// SIMATIC S7-200 project (STEP 7-Micro/WIN), CPU 224XP CN REL 02.01

SYMBOL_TABLE USUARIO1
SO               I0.3     // Sensor de Objetos (Detecta la pieza para iniciar la seleccion)
S_I              I0.4     // Sensor de fibra Optica (clasificacion de materiales)
SM               I0.5     // Sensor magnetico (clasificacion de materiales)
S1               I0.7     // Sensor de retorno del cilindro 1
S2               I1.0     // Sensor de retorno del cilindro 2
S3               I1.1     // Sensor de retorno del cilindro 3
SBB1             I1.3     // Pulsador de Marcha
SBB2             I1.2     // Pulsador de Paro
QS               I1.4     // Zeta de emergencia
SA               I1.5     // Selector rotatorio
am               Q0.0     // Motor
C_1              Q0.4     // cilindro neumatico 1
C_2              Q0.5     // cilindro neumatico 2
C_3              Q0.6     // cilindro neumatico 3
HL1              Q0.7     // Lampara de señalizacion amarilla
HL2              Q1.0     // Lampara de señalizacion verde
HL3              Q1.1     // Lampara de señalizacion roja
E0               M0.0     // Estado 0
E1               M0.1     // Estado 1
E2               M0.2     // Estado 2
E3               M0.3     // Estado 3
E4               M0.4     // Estado 4
E5               M0.5     // Estado 5
E6               M0.6     // Estado 6
E7               M0.7     // Estado 7
E8               M1.0     // Estado 8
E9               M1.1     // Estado 9
E10              M1.2     // Estado 10
E11              M1.3     // Estado 11
E12              M1.4     // Estado 12
E13              M1.5     // Estado 13
E14              M1.6     // Estado 14
EM               M1.7     // Variable para paro momentaneo
MOTOR            M2.0     // Variable para activacion o desactivacion del motor
E15              M2.1     // Estado 15
E16              M2.2     // Estado 16
C_c1             VD100
C_0              VD110
y_k              VD180
r_k              VD190
u_k              VD120
xh1_k_1          VD130
xh1_k            VD140
xh2_k_1          VD300
xh2_k            VD160
xh3_k_1          VD170
xh3_k            VD200
xp1_k            VD210
xp2_k            VD220
xp3_k            VD230
Ao               VD310
Bo               VD320
Co               VD330
Do               VD340
Eo               VD350
Fo               VD360
Go               VD370
Ho               VD380
Io               VD390
Jo               VD400
L1o              VD410
L2o              VD420
L3o              VD430
e_k              VD270
Ee               VD240
r_k_1            VD250
u_k_1            VD150
k1o              VD440
k2o              VD450
k3o              VD460
END_SYMBOL_TABLE

ORGANIZATION_BLOCK PRINCIPAL:OB1
TITLE=UNIDAD DE SELECCION
BEGIN
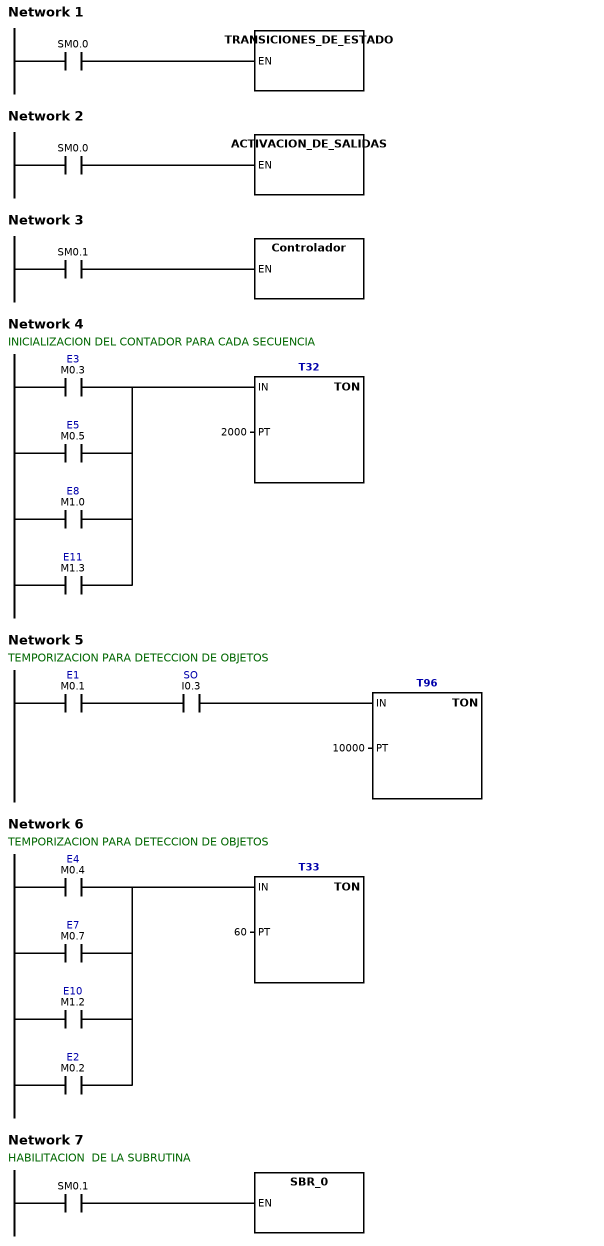
Network 1
LD     SM0.0
CALL   TRANSICIONES_DE_ESTADO:SBR1
Network 2
LD     SM0.0
CALL   ACTIVACION_DE_SALIDAS:SBR2
Network 3
LD     SM0.1
CALL   Controlador:SBR3
Network 4
// INICIALIZACION DEL CONTADOR PARA CADA SECUENCIA 
LD     E3:M0.3
O      E5:M0.5
O      E8:M1.0
O      E11:M1.3
TON    T32, 2000
Network 5
// TEMPORIZACION PARA DETECCION DE OBJETOS
LD     E1:M0.1
A      SO:I0.3
TON    T96, 10000
Network 6
// TEMPORIZACION PARA DETECCION DE OBJETOS
LD     E4:M0.4
O      E7:M0.7
O      E10:M1.2
O      E2:M0.2
TON    T33, 60
Network 7
// HABILITACION  DE LA SUBRUTINA
LD     SM0.1
CALL   SBR_0:SBR0
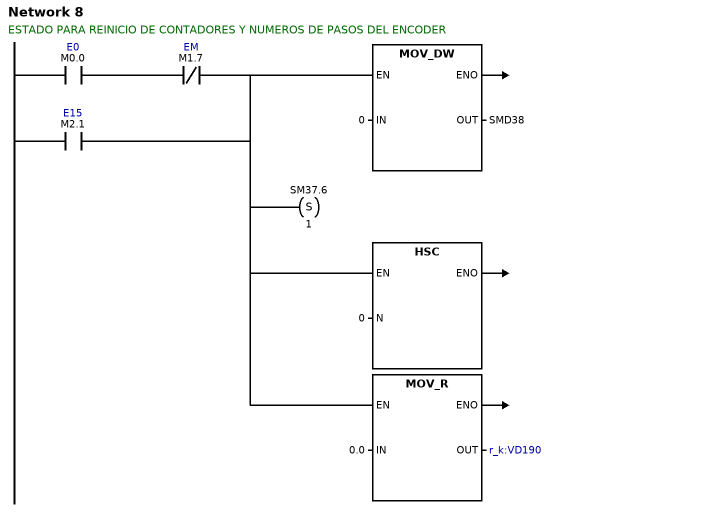
Network 8
// ESTADO PARA REINICIO DE CONTADORES Y NUMEROS DE PASOS DEL ENCODER
LD     E0:M0.0
AN     EM:M1.7
O      E15:M2.1
MOVD   0, SMD38
S      SM37.6, 1
HSC    0
MOVR   0.0, r_k:VD190
END_ORGANIZATION_BLOCK

SUBROUTINE_BLOCK SBR_0:SBR0
TITLE=COMENTARIOS DE LA SUBRUTINA
BEGIN
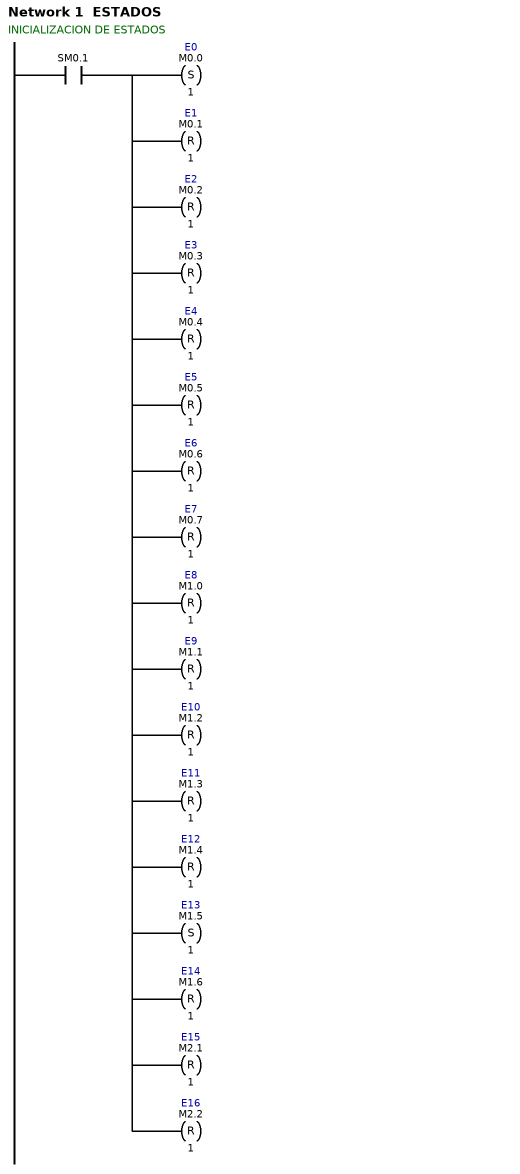
Network 1 // ESTADOS
// INICIALIZACION DE ESTADOS
LD     SM0.1
S      E0:M0.0, 1
R      E1:M0.1, 1
R      E2:M0.2, 1
R      E3:M0.3, 1
R      E4:M0.4, 1
R      E5:M0.5, 1
R      E6:M0.6, 1
R      E7:M0.7, 1
R      E8:M1.0, 1
R      E9:M1.1, 1
R      E10:M1.2, 1
R      E11:M1.3, 1
R      E12:M1.4, 1
S      E13:M1.5, 1
R      E14:M1.6, 1
R      E15:M2.1, 1
R      E16:M2.2, 1
END_SUBROUTINE_BLOCK

SUBROUTINE_BLOCK TRANSICIONES_DE_ESTADO:SBR1
TITLE=TRANSICIONES DE ESTADO
BEGIN
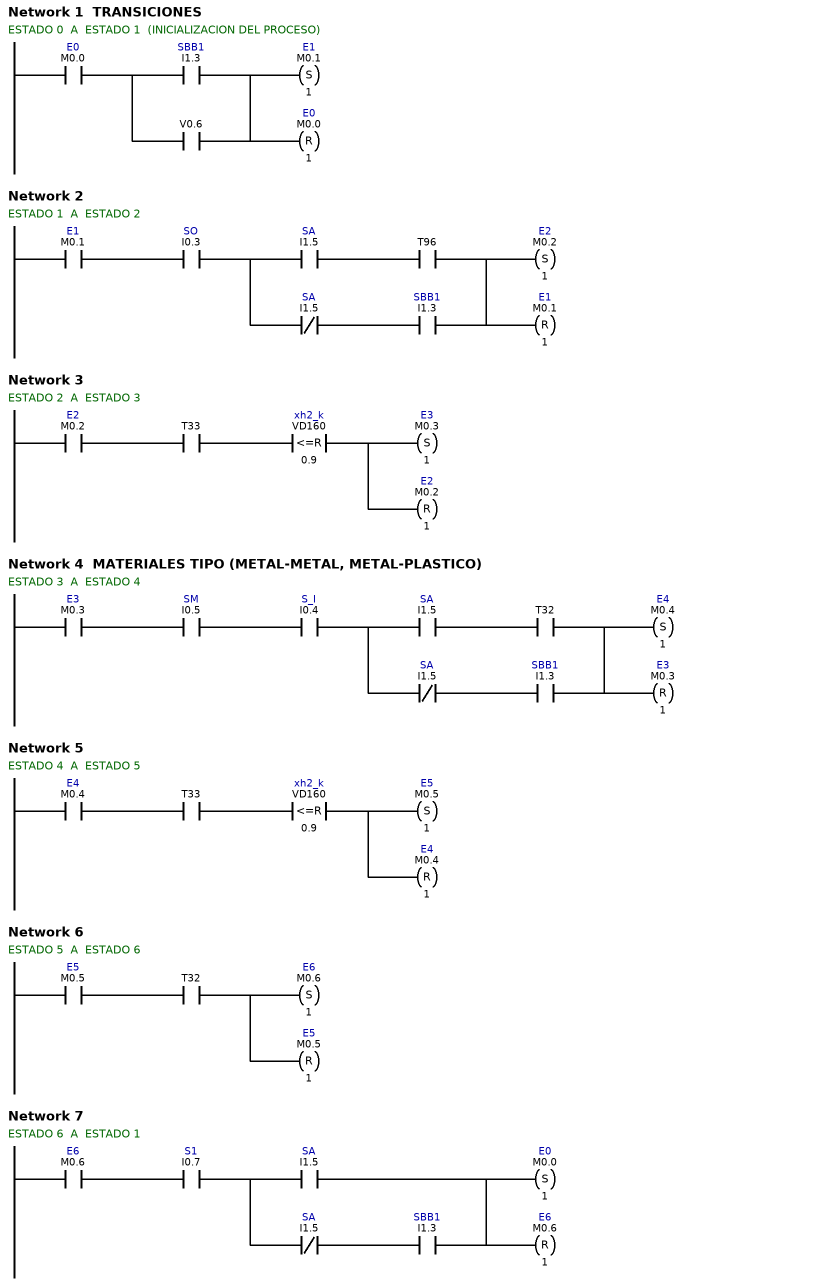
Network 1 // TRANSICIONES
// ESTADO 0  A  ESTADO 1  (INICIALIZACION DEL PROCESO)
LD     E0:M0.0
LD     SBB1:I1.3
O      V0.6
ALD
S      E1:M0.1, 1
R      E0:M0.0, 1
Network 2
// ESTADO 1  A  ESTADO 2 
LD     E1:M0.1
A      SO:I0.3
LD     SA:I1.5
A      T96
LDN    SA:I1.5
A      SBB1:I1.3
OLD
ALD
S      E2:M0.2, 1
R      E1:M0.1, 1
Network 3
// ESTADO 2  A  ESTADO 3
LD     E2:M0.2
A      T33
AR<=   xh2_k:VD160, 0.9
S      E3:M0.3, 1
R      E2:M0.2, 1
Network 4 // MATERIALES TIPO (METAL-METAL, METAL-PLASTICO)
// ESTADO 3  A  ESTADO 4
LD     E3:M0.3
A      SM:I0.5
A      S_I:I0.4
LD     SA:I1.5
A      T32
LDN    SA:I1.5
A      SBB1:I1.3
OLD
ALD
S      E4:M0.4, 1
R      E3:M0.3, 1
Network 5
// ESTADO 4  A  ESTADO 5
LD     E4:M0.4
A      T33
AR<=   xh2_k:VD160, 0.9
S      E5:M0.5, 1
R      E4:M0.4, 1
Network 6
// ESTADO 5  A  ESTADO 6
LD     E5:M0.5
A      T32
S      E6:M0.6, 1
R      E5:M0.5, 1
Network 7
// ESTADO 6  A  ESTADO 1
LD     E6:M0.6
A      S1:I0.7
LD     SA:I1.5
LDN    SA:I1.5
A      SBB1:I1.3
OLD
ALD
S      E0:M0.0, 1
R      E6:M0.6, 1
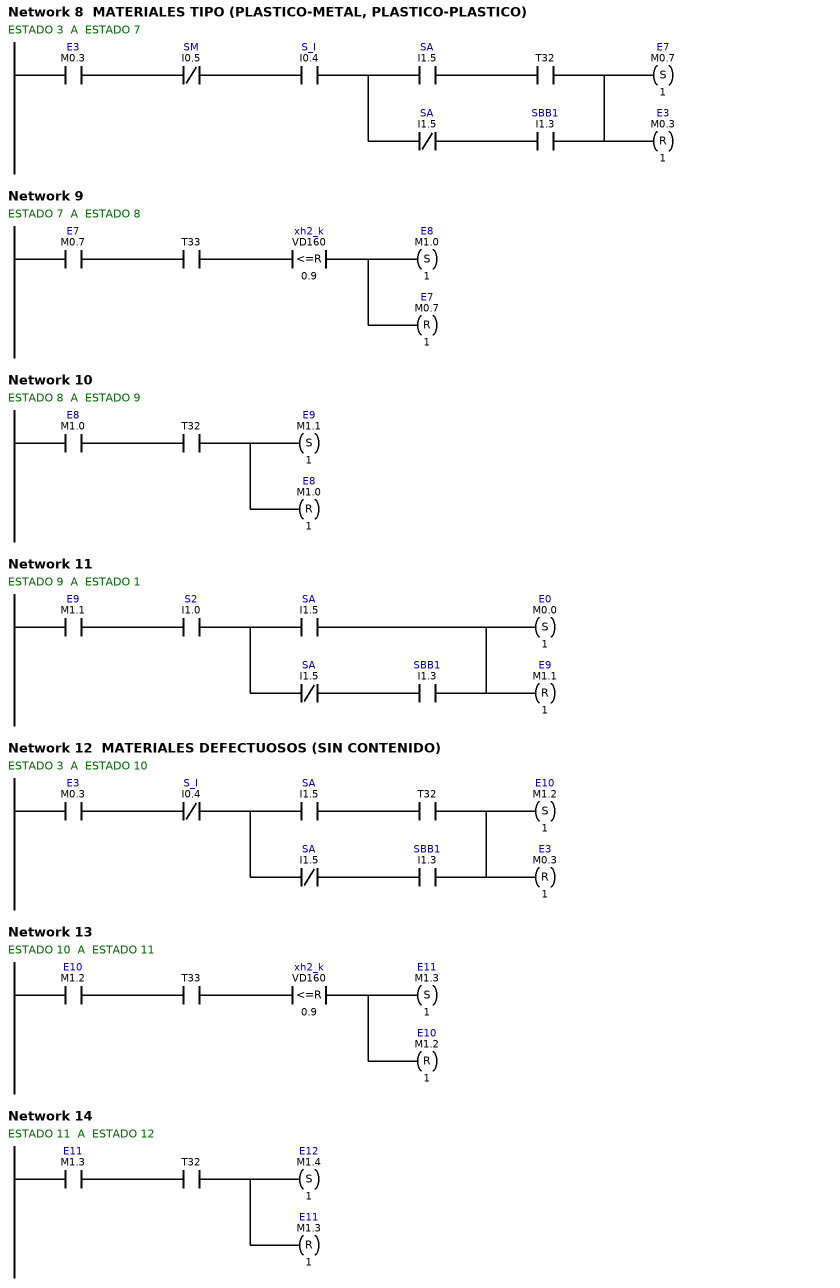
Network 8 // MATERIALES TIPO (PLASTICO-METAL, PLASTICO-PLASTICO)
// ESTADO 3  A  ESTADO 7
LD     E3:M0.3
AN     SM:I0.5
A      S_I:I0.4
LD     SA:I1.5
A      T32
LDN    SA:I1.5
A      SBB1:I1.3
OLD
ALD
S      E7:M0.7, 1
R      E3:M0.3, 1
Network 9
// ESTADO 7  A  ESTADO 8
LD     E7:M0.7
A      T33
AR<=   xh2_k:VD160, 0.9
S      E8:M1.0, 1
R      E7:M0.7, 1
Network 10
// ESTADO 8  A  ESTADO 9
LD     E8:M1.0
A      T32
S      E9:M1.1, 1
R      E8:M1.0, 1
Network 11
// ESTADO 9  A  ESTADO 1
LD     E9:M1.1
A      S2:I1.0
LD     SA:I1.5
LDN    SA:I1.5
A      SBB1:I1.3
OLD
ALD
S      E0:M0.0, 1
R      E9:M1.1, 1
Network 12 // MATERIALES DEFECTUOSOS (SIN CONTENIDO)
// ESTADO 3  A  ESTADO 10 
LD     E3:M0.3
AN     S_I:I0.4
LD     SA:I1.5
A      T32
LDN    SA:I1.5
A      SBB1:I1.3
OLD
ALD
S      E10:M1.2, 1
R      E3:M0.3, 1
Network 13
// ESTADO 10  A  ESTADO 11
LD     E10:M1.2
A      T33
AR<=   xh2_k:VD160, 0.9
S      E11:M1.3, 1
R      E10:M1.2, 1
Network 14
// ESTADO 11  A  ESTADO 12
LD     E11:M1.3
A      T32
S      E12:M1.4, 1
R      E11:M1.3, 1
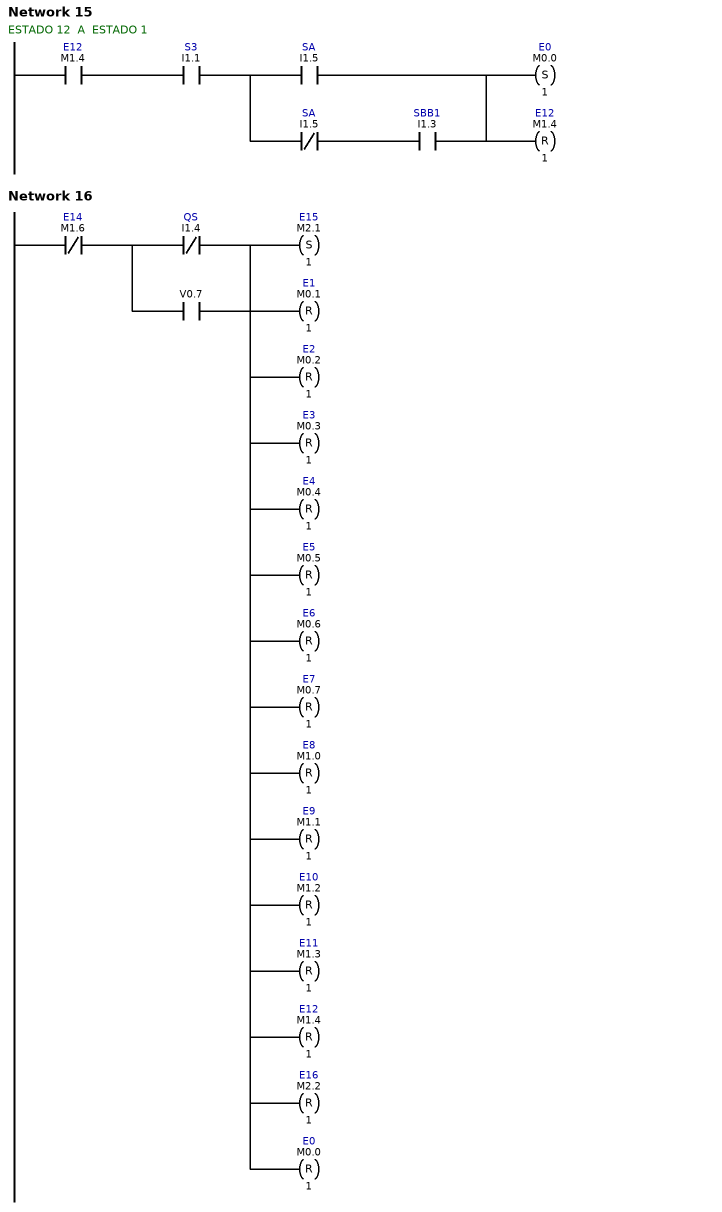
Network 15
// ESTADO 12  A  ESTADO 1
LD     E12:M1.4
A      S3:I1.1
LD     SA:I1.5
LDN    SA:I1.5
A      SBB1:I1.3
OLD
ALD
S      E0:M0.0, 1
R      E12:M1.4, 1
Network 16
LDN    E14:M1.6
LDN    QS:I1.4
O      V0.7
ALD
S      E15:M2.1, 1
R      E1:M0.1, 1
R      E2:M0.2, 1
R      E3:M0.3, 1
R      E4:M0.4, 1
R      E5:M0.5, 1
R      E6:M0.6, 1
R      E7:M0.7, 1
R      E8:M1.0, 1
R      E9:M1.1, 1
R      E10:M1.2, 1
R      E11:M1.3, 1
R      E12:M1.4, 1
R      E16:M2.2, 1
R      E0:M0.0, 1
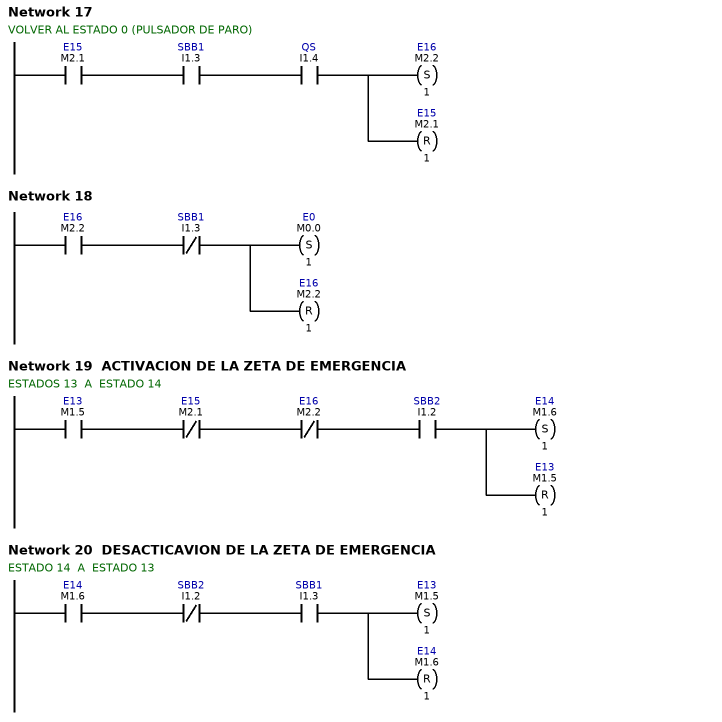
Network 17
// VOLVER AL ESTADO 0 (PULSADOR DE PARO)
LD     E15:M2.1
A      SBB1:I1.3
A      QS:I1.4
S      E16:M2.2, 1
R      E15:M2.1, 1
Network 18
LD     E16:M2.2
AN     SBB1:I1.3
S      E0:M0.0, 1
R      E16:M2.2, 1
Network 19 // ACTIVACION DE LA ZETA DE EMERGENCIA
// ESTADOS 13  A  ESTADO 14
LD     E13:M1.5
AN     E15:M2.1
AN     E16:M2.2
A      SBB2:I1.2
S      E14:M1.6, 1
R      E13:M1.5, 1
Network 20 // DESACTICAVION DE LA ZETA DE EMERGENCIA
// ESTADO 14  A  ESTADO 13
LD     E14:M1.6
AN     SBB2:I1.2
A      SBB1:I1.3
S      E13:M1.5, 1
R      E14:M1.6, 1
Network 21 // Título de segmento
// Comentario de segmento
END_SUBROUTINE_BLOCK

SUBROUTINE_BLOCK ACTIVACION_DE_SALIDAS:SBR2
TITLE=COMENTARIOS DE LA SUBRUTINA
BEGIN
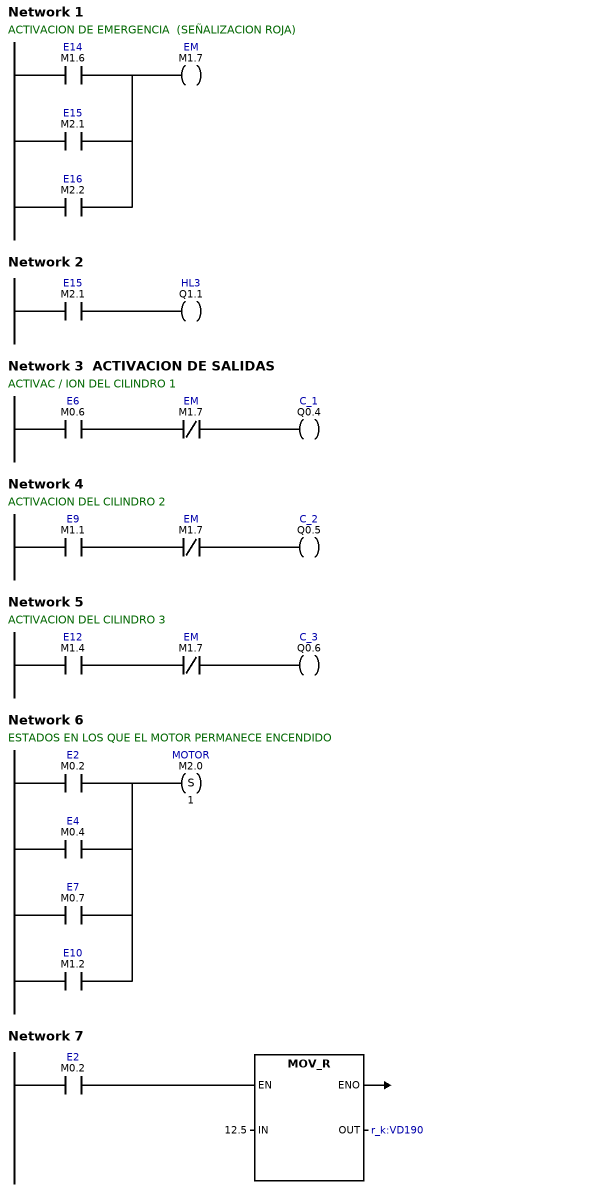
Network 1
// ACTIVACION DE EMERGENCIA  (SEÑALIZACION ROJA)
LD     E14:M1.6
O      E15:M2.1
O      E16:M2.2
=      EM:M1.7
Network 2
LD     E15:M2.1
=      HL3:Q1.1
Network 3 // ACTIVACION DE SALIDAS
// ACTIVAC
// ION DEL CILINDRO 1
LD     E6:M0.6
AN     EM:M1.7
=      C_1:Q0.4
Network 4
// ACTIVACION DEL CILINDRO 2
LD     E9:M1.1
AN     EM:M1.7
=      C_2:Q0.5
Network 5
// ACTIVACION DEL CILINDRO 3
LD     E12:M1.4
AN     EM:M1.7
=      C_3:Q0.6
Network 6
// ESTADOS EN LOS QUE EL MOTOR PERMANECE ENCENDIDO
LD     E2:M0.2
O      E4:M0.4
O      E7:M0.7
O      E10:M1.2
S      MOTOR:M2.0, 1
Network 7
LD     E2:M0.2
MOVR   12.5, r_k:VD190
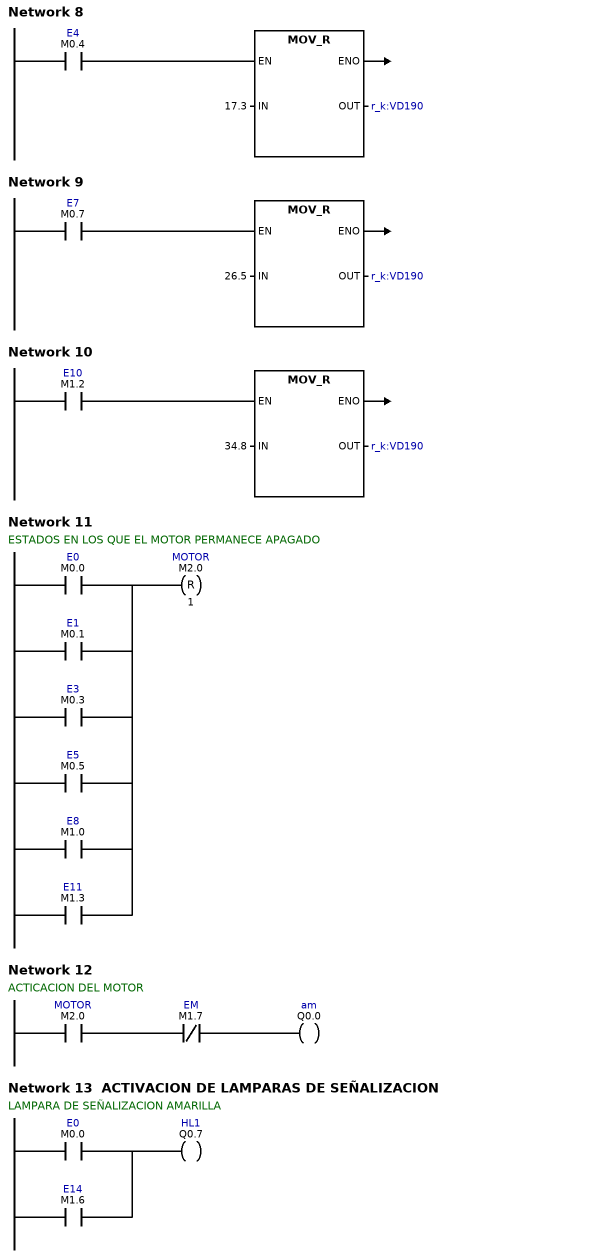
Network 8
LD     E4:M0.4
MOVR   17.3, r_k:VD190
Network 9
LD     E7:M0.7
MOVR   26.5, r_k:VD190
Network 10
LD     E10:M1.2
MOVR   34.8, r_k:VD190
Network 11
// ESTADOS EN LOS QUE EL MOTOR PERMANECE APAGADO
LD     E0:M0.0
O      E1:M0.1
O      E3:M0.3
O      E5:M0.5
O      E8:M1.0
O      E11:M1.3
R      MOTOR:M2.0, 1
Network 12
// ACTICACION DEL MOTOR
LD     MOTOR:M2.0
AN     EM:M1.7
=      am:Q0.0
Network 13 // ACTIVACION DE LAMPARAS DE SEÑALIZACION
// LAMPARA DE SEÑALIZACION AMARILLA
LD     E0:M0.0
O      E14:M1.6
=      HL1:Q0.7
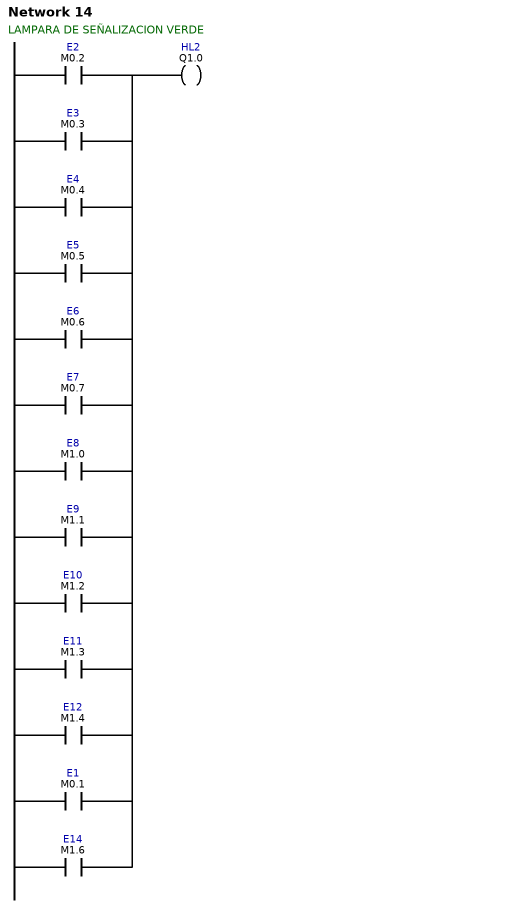
Network 14
// LAMPARA DE SEÑALIZACION VERDE
LD     E2:M0.2
O      E3:M0.3
O      E4:M0.4
O      E5:M0.5
O      E6:M0.6
O      E7:M0.7
O      E8:M1.0
O      E9:M1.1
O      E10:M1.2
O      E11:M1.3
O      E12:M1.4
O      E1:M0.1
O      E14:M1.6
=      HL2:Q1.0
Network 15 // Título de segmento
// Comentario de segmento
END_SUBROUTINE_BLOCK

SUBROUTINE_BLOCK Controlador:SBR3
TITLE=
BEGIN
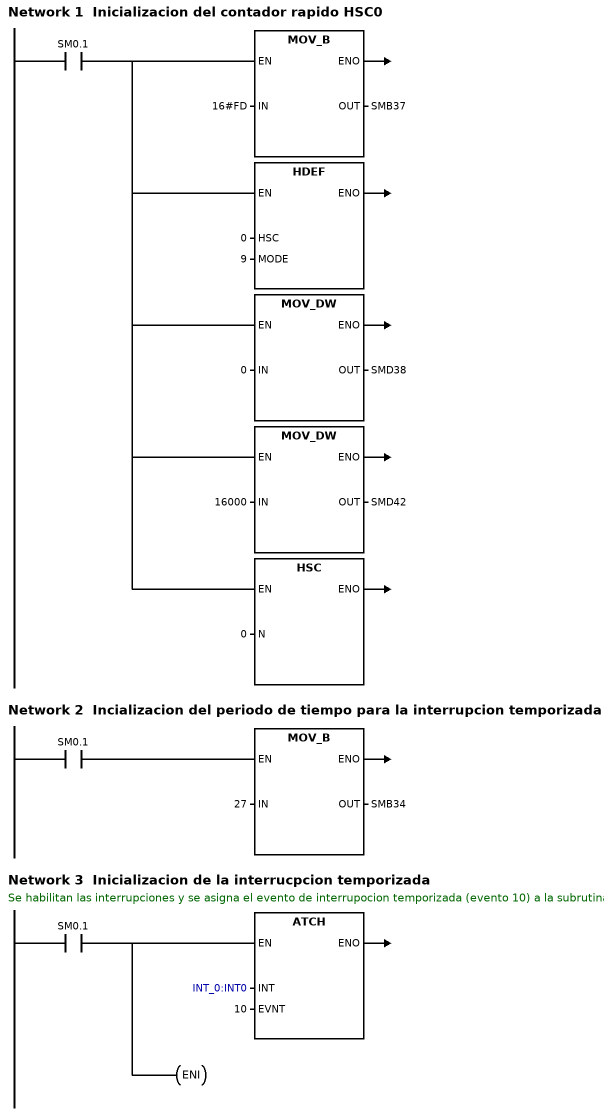
Network 1 // Inicializacion del contador rapido HSC0
LD     SM0.1
MOVB   16#FD, SMB37
HDEF   0, 9
MOVD   0, SMD38
MOVD   16000, SMD42
HSC    0
Network 2 // Incializacion del periodo de tiempo para la interrupcion temporizada
LD     SM0.1
MOVB   27, SMB34
Network 3 // Inicializacion de la interrucpcion temporizada
// Se habilitan las interrupciones y se asigna el evento de interrupocion temporizada (evento 10) a la subrutina de interrupcion INT_0
LD     SM0.1
ATCH   INT_0:INT0, 10
ENI
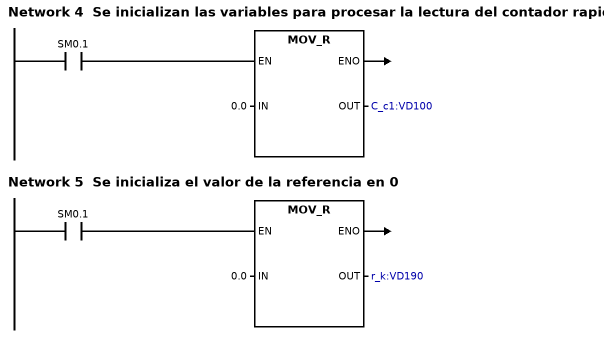
Network 4 // Se inicializan las variables para procesar la lectura del contador rapido HSC0
LD     SM0.1
MOVR   0.0, C_c1:VD100
Network 5 // Se inicializa el valor de la referencia en 0
LD     SM0.1
MOVR   0.0, r_k:VD190
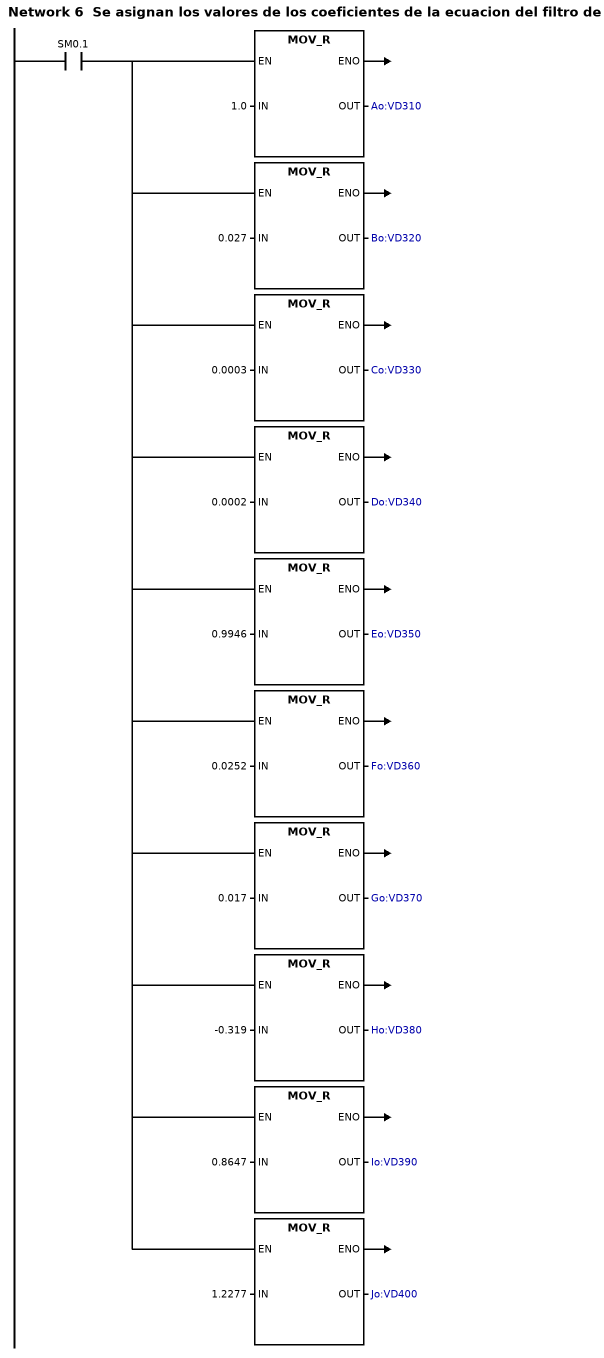
Network 6 // Se asignan los valores de los coeficientes de la ecuacion del filtro de KALMAN
LD     SM0.1
MOVR   1.0, Ao:VD310
MOVR   0.027, Bo:VD320
MOVR   0.0003, Co:VD330
MOVR   0.0002, Do:VD340
MOVR   0.9946, Eo:VD350
MOVR   0.0252, Fo:VD360
MOVR   0.017, Go:VD370
MOVR   -0.319, Ho:VD380
MOVR   0.8647, Io:VD390
MOVR   1.2277, Jo:VD400
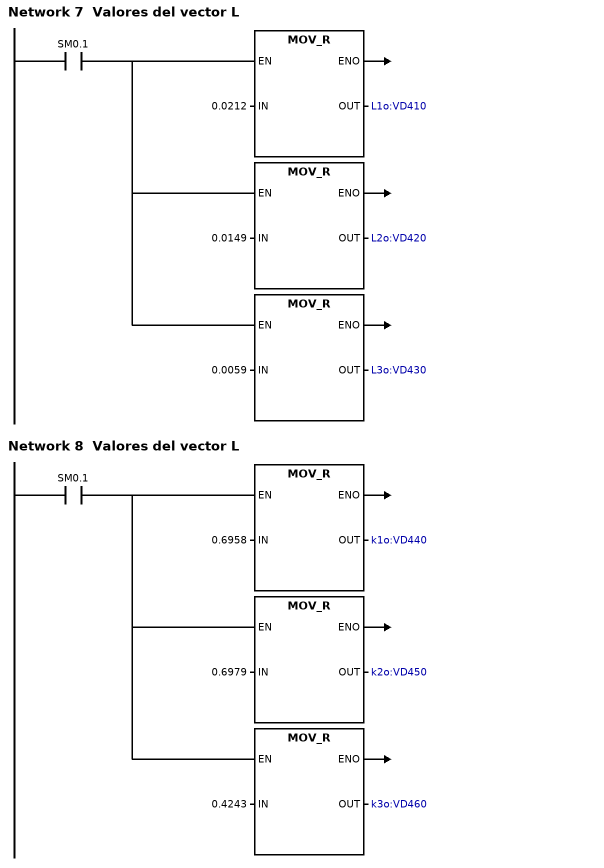
Network 7 // Valores del vector L
LD     SM0.1
MOVR   0.0212, L1o:VD410
MOVR   0.0149, L2o:VD420
MOVR   0.0059, L3o:VD430
Network 8 // Valores del vector L
LD     SM0.1
MOVR   0.6958, k1o:VD440
MOVR   0.6979, k2o:VD450
MOVR   0.4243, k3o:VD460
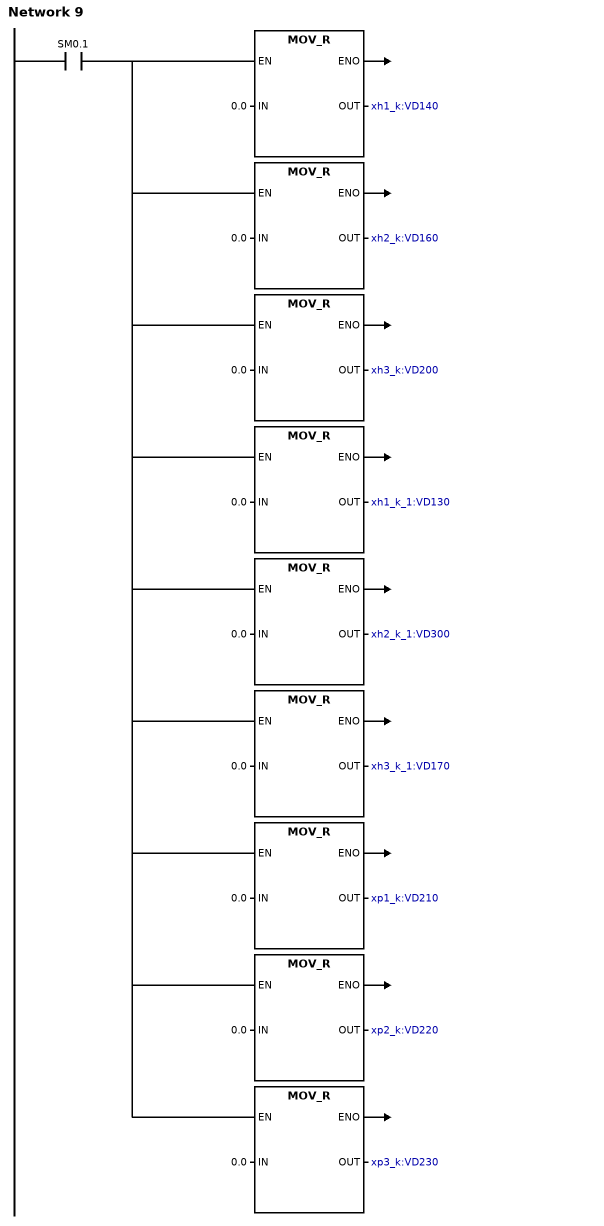
Network 9
LD     SM0.1
MOVR   0.0, xh1_k:VD140
MOVR   0.0, xh2_k:VD160
MOVR   0.0, xh3_k:VD200
MOVR   0.0, xh1_k_1:VD130
MOVR   0.0, xh2_k_1:VD300
MOVR   0.0, xh3_k_1:VD170
MOVR   0.0, xp1_k:VD210
MOVR   0.0, xp2_k:VD220
MOVR   0.0, xp3_k:VD230
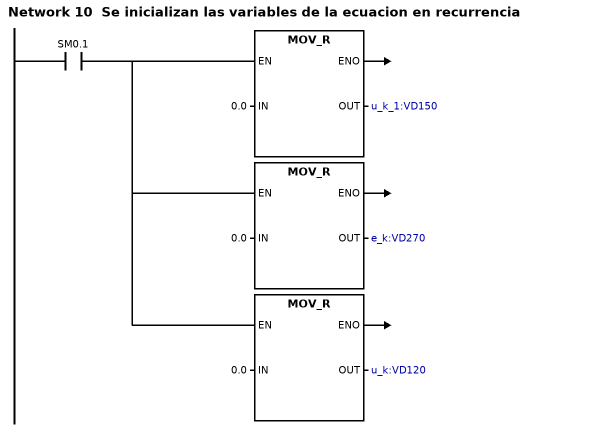
Network 10 // Se inicializan las variables de la ecuacion en recurrencia
LD     SM0.1
MOVR   0.0, u_k_1:VD150
MOVR   0.0, e_k:VD270
MOVR   0.0, u_k:VD120
END_SUBROUTINE_BLOCK

INTERRUPT_BLOCK INT_0:INT0
TITLE=COMENTARIOS DE LA RUTINA DE INTERRUPCIÓN
BEGIN
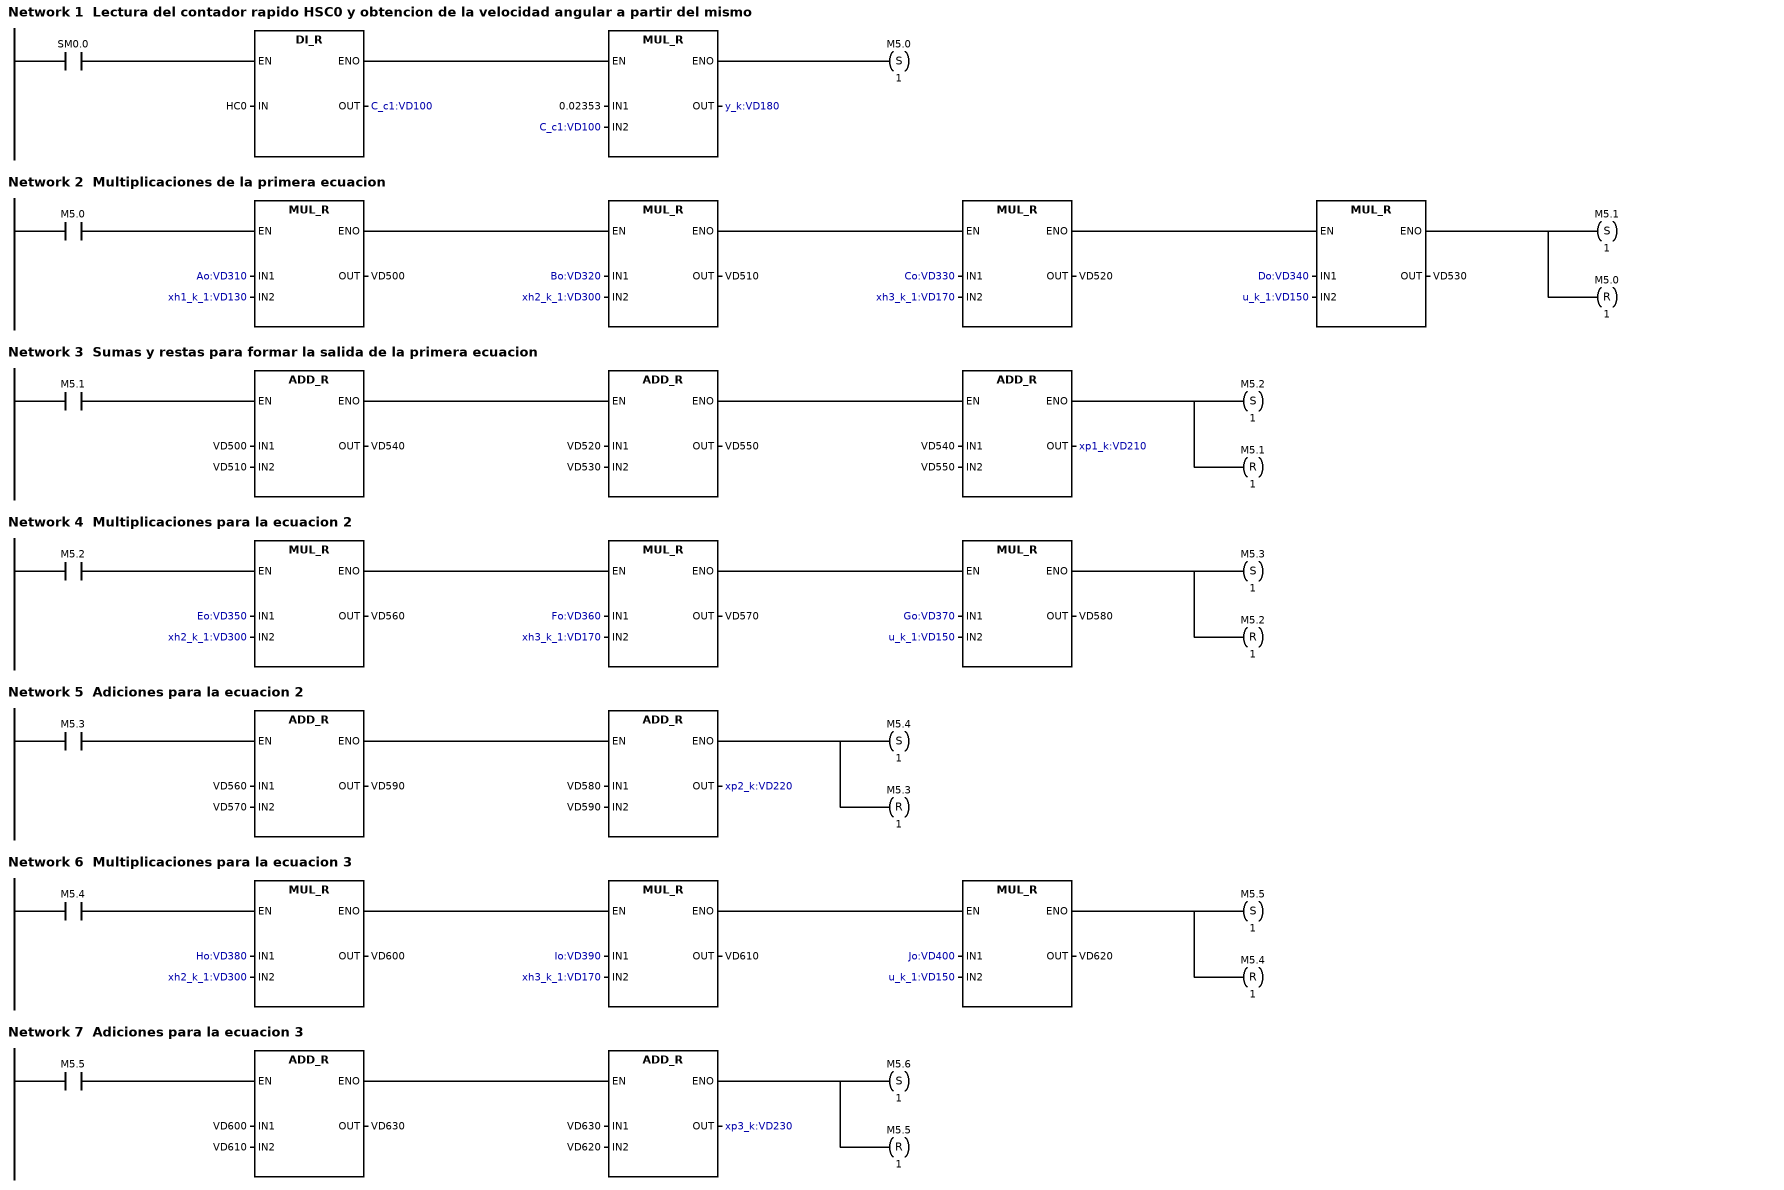
Network 1 // Lectura del contador rapido HSC0 y obtencion de la velocidad angular a partir del mismo
LD     SM0.0
DTR    HC0, C_c1:VD100
AENO
MOVR   0.02353, y_k:VD180
AENO
*R     C_c1:VD100, y_k:VD180
AENO
S      M5.0, 1
Network 2 // Multiplicaciones de la primera ecuacion 
LD     M5.0
MOVR   Ao:VD310, VD500
AENO
*R     xh1_k_1:VD130, VD500
AENO
MOVR   Bo:VD320, VD510
AENO
*R     xh2_k_1:VD300, VD510
AENO
MOVR   Co:VD330, VD520
AENO
*R     xh3_k_1:VD170, VD520
AENO
MOVR   Do:VD340, VD530
AENO
*R     u_k_1:VD150, VD530
AENO
S      M5.1, 1
R      M5.0, 1
Network 3 // Sumas y restas para formar la salida de la primera ecuacion
LD     M5.1
MOVR   VD500, VD540
AENO
+R     VD510, VD540
AENO
MOVR   VD520, VD550
AENO
+R     VD530, VD550
AENO
MOVR   VD540, xp1_k:VD210
AENO
+R     VD550, xp1_k:VD210
AENO
S      M5.2, 1
R      M5.1, 1
Network 4 // Multiplicaciones para la ecuacion 2
LD     M5.2
MOVR   Eo:VD350, VD560
AENO
*R     xh2_k_1:VD300, VD560
AENO
MOVR   Fo:VD360, VD570
AENO
*R     xh3_k_1:VD170, VD570
AENO
MOVR   Go:VD370, VD580
AENO
*R     u_k_1:VD150, VD580
AENO
S      M5.3, 1
R      M5.2, 1
Network 5 // Adiciones para la ecuacion 2
LD     M5.3
MOVR   VD560, VD590
AENO
+R     VD570, VD590
AENO
MOVR   VD580, xp2_k:VD220
AENO
+R     VD590, xp2_k:VD220
AENO
S      M5.4, 1
R      M5.3, 1
Network 6 // Multiplicaciones para la ecuacion 3
LD     M5.4
MOVR   Ho:VD380, VD600
AENO
*R     xh2_k_1:VD300, VD600
AENO
MOVR   Io:VD390, VD610
AENO
*R     xh3_k_1:VD170, VD610
AENO
MOVR   Jo:VD400, VD620
AENO
*R     u_k_1:VD150, VD620
AENO
S      M5.5, 1
R      M5.4, 1
Network 7 // Adiciones para la ecuacion 3
LD     M5.5
MOVR   VD600, VD630
AENO
+R     VD610, VD630
AENO
MOVR   VD630, xp3_k:VD230
AENO
+R     VD620, xp3_k:VD230
AENO
S      M5.6, 1
R      M5.5, 1
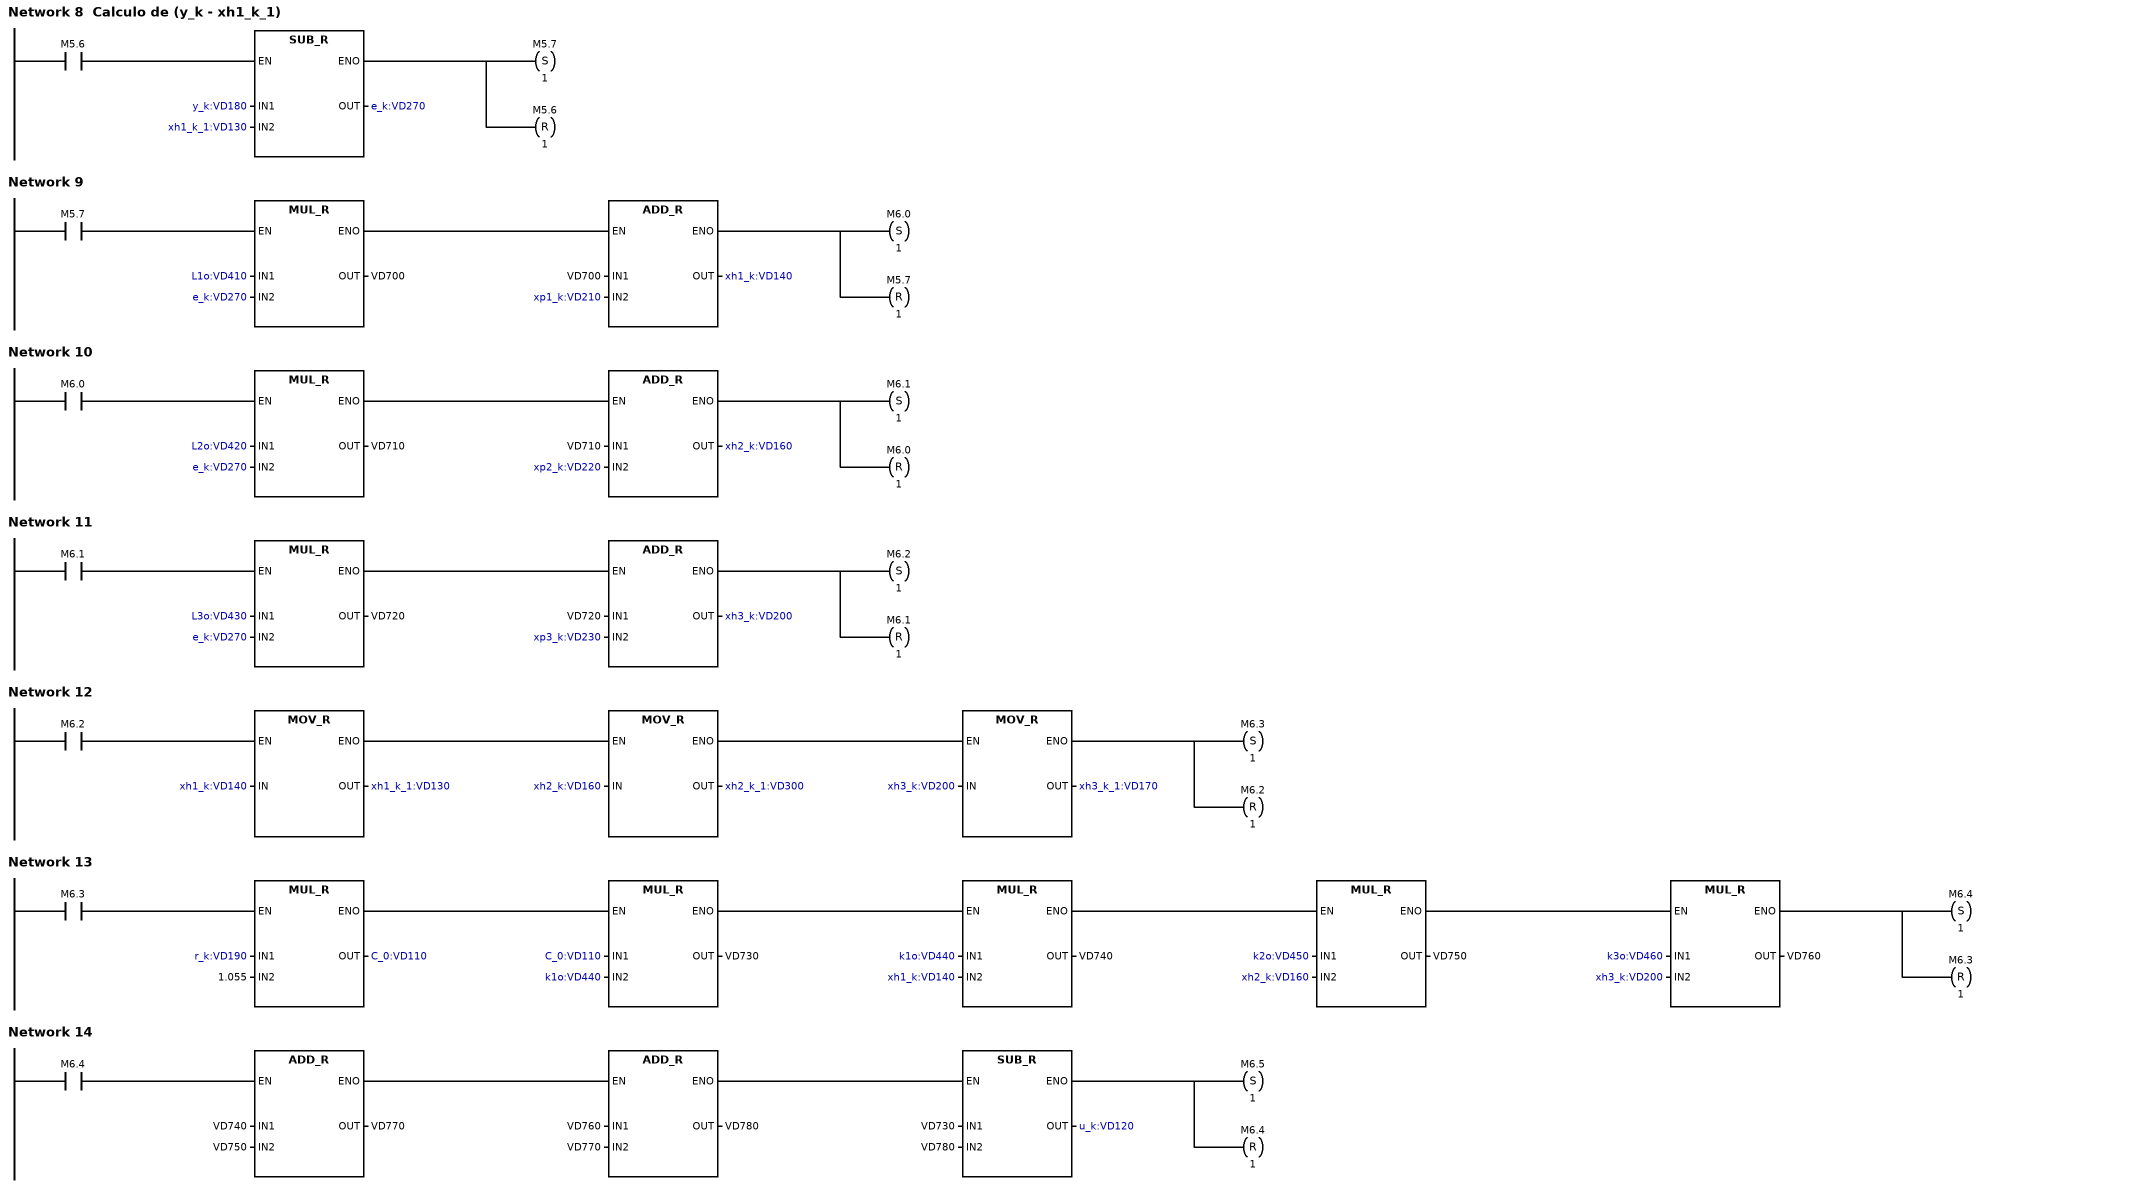
Network 8 // Calculo de (y_k - xh1_k_1)
LD     M5.6
MOVR   y_k:VD180, e_k:VD270
AENO
-R     xh1_k_1:VD130, e_k:VD270
AENO
S      M5.7, 1
R      M5.6, 1
Network 9
LD     M5.7
MOVR   L1o:VD410, VD700
AENO
*R     e_k:VD270, VD700
AENO
MOVR   VD700, xh1_k:VD140
AENO
+R     xp1_k:VD210, xh1_k:VD140
AENO
S      M6.0, 1
R      M5.7, 1
Network 10
LD     M6.0
MOVR   L2o:VD420, VD710
AENO
*R     e_k:VD270, VD710
AENO
MOVR   VD710, xh2_k:VD160
AENO
+R     xp2_k:VD220, xh2_k:VD160
AENO
S      M6.1, 1
R      M6.0, 1
Network 11
LD     M6.1
MOVR   L3o:VD430, VD720
AENO
*R     e_k:VD270, VD720
AENO
MOVR   VD720, xh3_k:VD200
AENO
+R     xp3_k:VD230, xh3_k:VD200
AENO
S      M6.2, 1
R      M6.1, 1
Network 12
LD     M6.2
MOVR   xh1_k:VD140, xh1_k_1:VD130
AENO
MOVR   xh2_k:VD160, xh2_k_1:VD300
AENO
MOVR   xh3_k:VD200, xh3_k_1:VD170
AENO
S      M6.3, 1
R      M6.2, 1
Network 13
LD     M6.3
MOVR   r_k:VD190, C_0:VD110
AENO
*R     1.055, C_0:VD110
AENO
MOVR   C_0:VD110, VD730
AENO
*R     k1o:VD440, VD730
AENO
MOVR   k1o:VD440, VD740
AENO
*R     xh1_k:VD140, VD740
AENO
MOVR   k2o:VD450, VD750
AENO
*R     xh2_k:VD160, VD750
AENO
MOVR   k3o:VD460, VD760
AENO
*R     xh3_k:VD200, VD760
AENO
S      M6.4, 1
R      M6.3, 1
Network 14
LD     M6.4
MOVR   VD740, VD770
AENO
+R     VD750, VD770
AENO
MOVR   VD760, VD780
AENO
+R     VD770, VD780
AENO
MOVR   VD730, u_k:VD120
AENO
-R     VD780, u_k:VD120
AENO
S      M6.5, 1
R      M6.4, 1
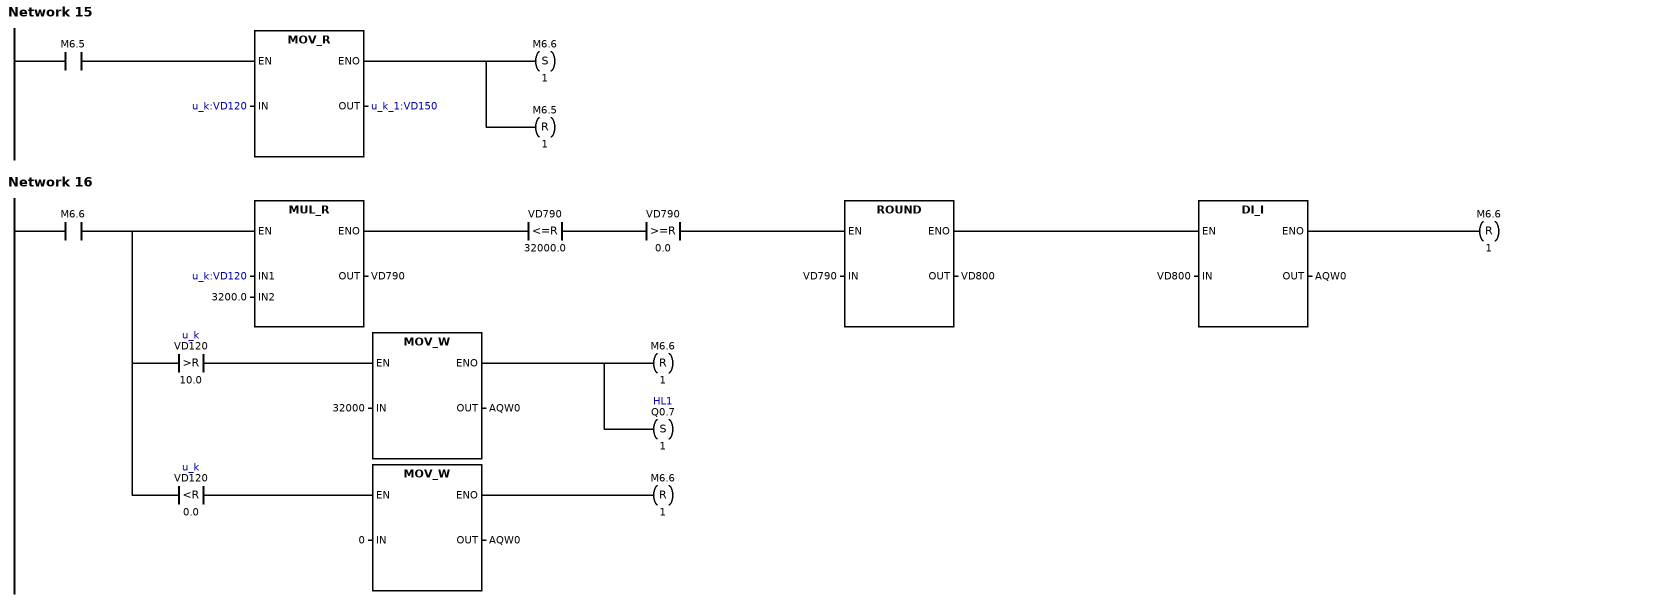
Network 15
LD     M6.5
MOVR   u_k:VD120, u_k_1:VD150
AENO
S      M6.6, 1
R      M6.5, 1
Network 16
LD     M6.6
LPS
MOVR   u_k:VD120, VD790
AENO
*R     3200.0, VD790
AENO
AR<=   VD790, 32000.0
AR>=   VD790, 0.0
ROUND  VD790, VD800
AENO
DTI    VD800, AQW0
AENO
R      M6.6, 1
LRD
AR>    u_k:VD120, 10.0
MOVW   32000, AQW0
AENO
R      M6.6, 1
S      HL1:Q0.7, 1
LPP
AR<    u_k:VD120, 0.0
MOVW   0, AQW0
AENO
R      M6.6, 1
Network 17 // Título de segmento
// Comentario de segmento
END_INTERRUPT_BLOCK
